// TIA Portal V21 export
// export: Created 2026-11-21T13:24:04.9288632Z, ExportSetting WithDefaults, DisplayName Totally Integrated Automation Portal, DisplayVersion V21, DisplayName STEP 7 Professional, DisplayVersion V21, DisplayName STEP 7 Safety, DisplayVersion V21, DisplayName Tech WebApplication, DisplayVersion V21, DisplayName WinCC Basic/Comfort/Advanced, DisplayVersion V21, DisplayName WinCC Unified, DisplayVersion V21
VAR_GLOBAL   // PLC tag table "Standard"
   Running AT %M10.0 : Bool;   // What the safety program released, for the standard program
END_VAR
